Fanuc KAREL source: KD00043.KL

PROGRAM KD00043
%NOLOCKGROUP
VAR
  I: INTEGER
  J: INTEGER
  B: BOOLEAN
  R: REAL
  S: STRING[80]
  C: COMMON_ASSOC
BEGIN
  I = 1
END KD00043
